// TIA Portal V19 export
FUNCTION_BLOCK "AI"   // FB8, LAD
{ S7_Optimized_Access := 'TRUE' }
// stored: MemoryReserve 100, SetENOAutomatically false
   VAR_INPUT
      RAW_MIN : Int;
      RAW_MAX : Int;
      SCALE_MIN : Real;
      SCALE_MAX : Real;
      HH_SP : Real;
      HSP : Real;
      LL_SP : Real;
      LSP : Real;
      ALM_WT : Time := T#10S;
      INPUT : Int;
   END_VAR
   VAR_OUTPUT
      FAULT : Bool;
      HH_ALM : Bool;
      H_ALM : Bool;
      LL_ALM : Bool;
      L_ALM : Bool;
      SCALE_OUT : Real;
   END_VAR
   VAR
      AI : "SCALING";
      MAX_VALUE : Int;
      HH_TIME { S7_SetPoint := 'True'} : TON_TIME;
      H_TIME { S7_SetPoint := 'True'} : TON_TIME;
      LL_TIME { S7_SetPoint := 'True'} : TON_TIME;
      L_TIME { S7_SetPoint := 'True'} : TON_TIME;
   END_VAR
BEGIN

REGION Network 2 (SCL)

   IF #INPUT < -100 OR #INPUT > 27648 THEN
       #FAULT := 1;
   ELSE
       #FAULT := 0;
   END_IF;
   IF NOT #FAULT THEN
       #AI(RAW_MIN := #RAW_MIN,
           RAW_MAX := #RAW_MAX,
           INPUT := #INPUT,
           SCALE_MIN := #SCALE_MIN,
           SCALE_MAX := #SCALE_MAX,
           SCALE_OUT => #SCALE_OUT);
   ELSE
       #SCALE_OUT := 0.0;

   END_IF;
END_REGION

REGION Network 3
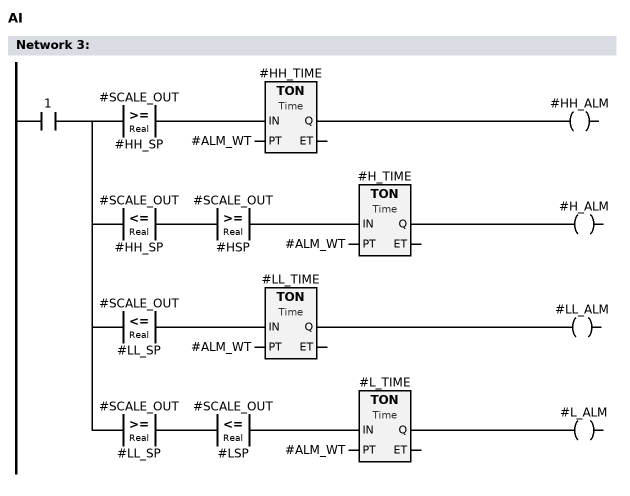
   RUNG wire#powerrail
      Contact( 1 )
      wire#w1
      { S7_Templates := "SrcType := Real" } GE_Contact(in1 := #SCALE_OUT, in2 := #HH_SP)
      { S7_Templates := "time_type := Time" } #HH_TIME.TON(pt := #ALM_WT, et =>)
      Coil( #HH_ALM )
   END_RUNG
   RUNG wire#w1
      { S7_Templates := "SrcType := Real" } LE_Contact(in1 := #SCALE_OUT, in2 := #HH_SP)
      { S7_Templates := "SrcType := Real" } GE_Contact(in1 := #SCALE_OUT, in2 := #HSP)
      { S7_Templates := "time_type := Time" } #H_TIME.TON(pt := #ALM_WT, et =>)
      Coil( #H_ALM )
   END_RUNG
   RUNG wire#w1
      { S7_Templates := "SrcType := Real" } LE_Contact(in1 := #SCALE_OUT, in2 := #LL_SP)
      { S7_Templates := "time_type := Time" } #LL_TIME.TON(pt := #ALM_WT, et =>)
      Coil( #LL_ALM )
   END_RUNG
   RUNG wire#w1
      { S7_Templates := "SrcType := Real" } GE_Contact(in1 := #SCALE_OUT, in2 := #LL_SP)
      { S7_Templates := "SrcType := Real" } LE_Contact(in1 := #SCALE_OUT, in2 := #LSP)
      { S7_Templates := "time_type := Time" } #L_TIME.TON(pt := #ALM_WT, et =>)
      Coil( #L_ALM )
   END_RUNG
   // the same network as SCL:
   #HH_TIME(IN := 1 AND (#SCALE_OUT >= #HH_SP), PT := #ALM_WT);   // TON
   #HH_ALM := #HH_TIME.Q;
   #H_TIME(IN := 1 AND (#SCALE_OUT <= #HH_SP) AND (#SCALE_OUT >= #HSP), PT := #ALM_WT);   // TON
   #H_ALM := #H_TIME.Q;
   #LL_TIME(IN := 1 AND (#SCALE_OUT <= #LL_SP), PT := #ALM_WT);   // TON
   #LL_ALM := #LL_TIME.Q;
   #L_TIME(IN := 1 AND (#SCALE_OUT >= #LL_SP) AND (#SCALE_OUT <= #LSP), PT := #ALM_WT);   // TON
   #L_ALM := #L_TIME.Q;
END_REGION
END_FUNCTION_BLOCK
